(* ================================================================= *)
(*  ST_InfeedSensors                                                  *)
(*  入料位置检测结构体 - 三段光电+去抖确认+参数                         *)
(*  版本: V1.0.0  日期: 2026-05-30                                    *)
(*  来源: SysLib/types/                                               *)
(*  复用: 工站输送机入料检测/多段光电位置确认                          *)
(*  引用: FB_1014_StationConveyor V2.0.0 改用VAR_IN_OUT引用           *)
(*                                                                    *)
(*  设计原则:                                                         *)
(*    - 原始传感器输入+去抖确认输出+参数同构                           *)
(*    - AllConfirmed由FB计算: StartConfirmed AND Pos1Confirmed         *)
(*      AND Pos2Confirmed                                             *)
(*    - DebounceMs统一配置三段光电去抖延时                             *)
(* ================================================================= *)

TYPE ST_InfeedSensors :
STRUCT
    // === Raw sensor inputs (OB1写入, FB读取) ===
    InfeedStart     : BOOL := FALSE;   // 入料开始光电 (入口检测)
    InfeedPos1      : BOOL := FALSE;   // 入料到位光电1 (粗定位)
    InfeedPos2      : BOOL := FALSE;   // 入料到位光电2 (精定位)

    // === Confirmed outputs (FB写入, 去抖后) ===
    StartConfirmed  : BOOL := FALSE;   // 入料开始确认
    Pos1Confirmed   : BOOL := FALSE;   // 到位1确认
    Pos2Confirmed   : BOOL := FALSE;   // 到位2确认
    AllConfirmed    : BOOL := FALSE;   // 三光电全部确认

    // === Parameter ===
    DebounceMs      : DINT := 200;     // 去抖延时 (ms), 50~2000
END_STRUCT
END_TYPE
